// FB MON state codes.
{attribute 'qualified_only'}
{attribute 'to_string'}
TYPE
E_SafeMonState :
(
    Undefined := 0,
    Run := 1,
    Stop := 2,
    Safe := 3,
    Error := 4,
    Reset := 5,
    Start := 6,
    ErrorDelay := 7,
    DelayOut := 8,
    FuncTest := 9
) BYTE;
END_TYPE

(* stored: Version 1.1.0.1
   DUT E_SafeMonState: Id {4195e8ba-862d-57bc-8b6f-9947275b3924} *)
